FUNCTION_BLOCK DLG_CTRL (* Ablaufsteuerung eines VT-Dialogs (MessageBox) *)
  (* Standard: 61499-2; Description: Copyright (c) 2026 Meisterschulen am Ostbahnhof This program and the accompanying materials are made available under the terms of the Eclipse Public License 2.0 which is available at https://www.eclipse.org/legal/epl-2.0/ SPDX-License-Identifier: EPL-2.0 *)
  (* Version 1.0, 2026-11-17, Franz Höpfinger, Meisterschulen am Ostbahnhof, initial API and implementation and/or initial documentation *)
  PACKAGE isobus::UT::dialog;
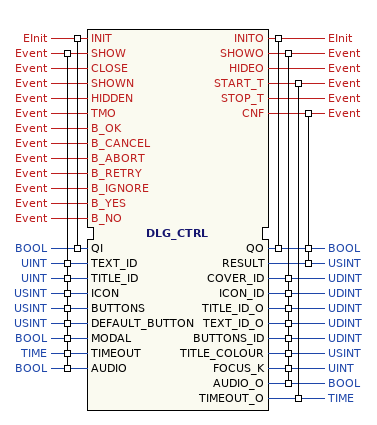
  EVENT_INPUT
    INIT : EInit WITH QI; (* Initialisierung *)
    SHOW WITH TEXT_ID, TITLE_ID, ICON, BUTTONS, DEFAULT_BUTTON, MODAL, TIMEOUT, AUDIO; (* Dialog zeigen *)
    CLOSE; (* Dialog vom Programm schliessen *)
    SHOWN; (* Anzeige-Kette fertig *)
    HIDDEN; (* Ausblenden fertig *)
    TMO; (* Zeit abgelaufen *)
    B_OK; (* Button OK losgelassen *)
    B_CANCEL; (* Button Cancel losgelassen *)
    B_ABORT; (* Button Abort losgelassen *)
    B_RETRY; (* Button Retry losgelassen *)
    B_IGNORE; (* Button Ignore losgelassen *)
    B_YES; (* Button Yes losgelassen *)
    B_NO; (* Button No losgelassen *)
  END_EVENT
  EVENT_OUTPUT
    INITO : EInit WITH QO; (* Initialisierung fertig *)
    SHOWO WITH COVER_ID, ICON_ID, TITLE_ID_O, TEXT_ID_O, BUTTONS_ID, TITLE_COLOUR, FOCUS_K, AUDIO_O; (* Anzeige-Kette starten *)
    HIDEO; (* Dialog ausblenden *)
    START_T WITH TIMEOUT_O; (* Timeout starten *)
    STOP_T; (* Timeout stoppen *)
    CNF WITH QO, RESULT; (* Dialog beendet *)
  END_EVENT
  VAR_INPUT
    QI : BOOL := TRUE; (* Freigabe *)
    TEXT_ID : UINT := UINT#65535; (* OutputString Meldungstext *)
    TITLE_ID : UINT := UINT#65535; (* OutputString Titel, NULL = Standard je Icon *)
    ICON : USINT := USINT#1; (* DLG_ICON_* *)
    BUTTONS : USINT := USINT#1; (* DLG_BTN_* *)
    DEFAULT_BUTTON : USINT := USINT#1; (* Fokus auf Taste 1..3 *)
    MODAL : BOOL := FALSE; (* Maske abdecken *)
    TIMEOUT : TIME := T#0s; (* T#0s = kein Timeout *)
    AUDIO : BOOL := FALSE; (* Ton beim Oeffnen *)
  END_VAR
  VAR_OUTPUT
    QO : BOOL; (* Qualitaet *)
    RESULT : USINT; (* DLG_RES_* *)
    COVER_ID : UDINT; (* Ziel ObjectPointer_Dlg_Cover *)
    ICON_ID : UDINT; (* Ziel ObjectPointer_Dlg_Icon *)
    TITLE_ID_O : UDINT; (* Ziel ObjectPointer_Dlg_Title *)
    TEXT_ID_O : UDINT; (* Ziel ObjectPointer_Dlg_Text *)
    BUTTONS_ID : UDINT; (* Ziel ObjectPointer_Dlg_Buttons *)
    TITLE_COLOUR : USINT; (* VT-Farbindex Titelzeile *)
    FOCUS_K : UINT; (* Fokus-Button 0..6, 7 = keiner *)
    AUDIO_O : BOOL; (* Ton ja/nein *)
    TIMEOUT_O : TIME; (* Timeout *)
  END_VAR
  VAR
    xPendingShow : BOOL; (* neues SHOW wartet *)
    xPendingClose : BOOL; (* Schliessen wartet *)
  END_VAR
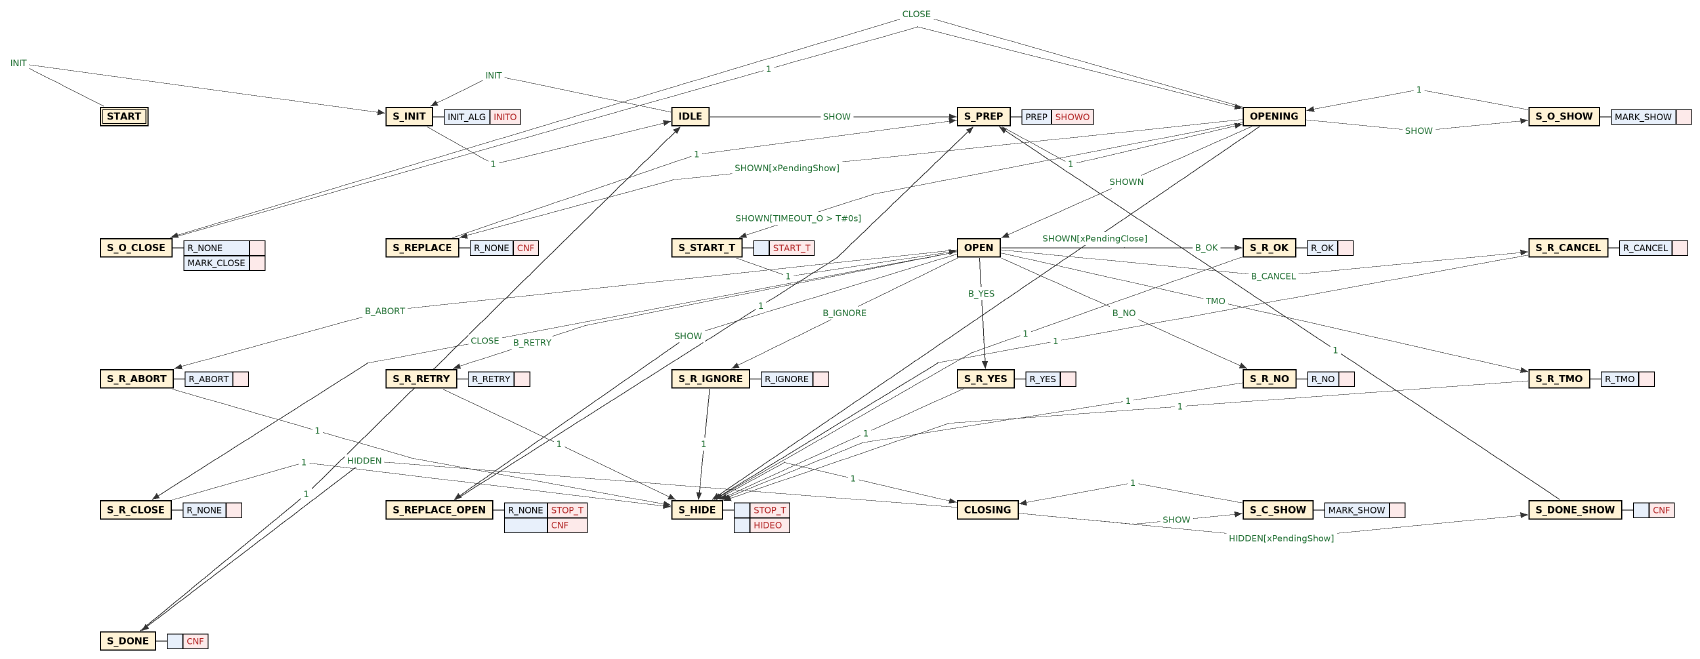
  EC_STATES
    START; (* Initial State *)
    S_INIT : INIT_ALG -> INITO;
    IDLE; (* kein Dialog offen *)
    S_PREP : PREP -> SHOWO; (* Anzeige-Kette starten *)
    OPENING; (* Anzeige-Kette laeuft *)
    S_O_SHOW : MARK_SHOW;
    S_O_CLOSE : R_NONE, MARK_CLOSE;
    S_REPLACE : R_NONE -> CNF; (* alter Dialog ersetzt *)
    S_START_T : -> START_T;
    OPEN; (* Dialog sichtbar *)
    S_R_OK : R_OK;
    S_R_CANCEL : R_CANCEL;
    S_R_ABORT : R_ABORT;
    S_R_RETRY : R_RETRY;
    S_R_IGNORE : R_IGNORE;
    S_R_YES : R_YES;
    S_R_NO : R_NO;
    S_R_TMO : R_TMO;
    S_R_CLOSE : R_NONE;
    S_REPLACE_OPEN : R_NONE -> STOP_T, -> CNF; (* neues SHOW waehrend offen *)
    S_HIDE : -> STOP_T, -> HIDEO;
    CLOSING; (* Ausblenden laeuft *)
    S_C_SHOW : MARK_SHOW;
    S_DONE_SHOW : -> CNF;
    S_DONE : -> CNF;
  END_STATES
  EC_TRANSITIONS
    START TO S_INIT := INIT;
    S_INIT TO IDLE := 1;
    IDLE TO S_INIT := INIT;
    IDLE TO S_PREP := SHOW;
    S_PREP TO OPENING := 1;
    OPENING TO S_HIDE := SHOWN[xPendingClose];
    OPENING TO S_REPLACE := SHOWN[xPendingShow];
    OPENING TO S_START_T := SHOWN[TIMEOUT_O > T#0s];
    OPENING TO OPEN := SHOWN;
    OPENING TO S_O_SHOW := SHOW;
    OPENING TO S_O_CLOSE := CLOSE;
    S_O_SHOW TO OPENING := 1;
    S_O_CLOSE TO OPENING := 1;
    S_REPLACE TO S_PREP := 1;
    S_START_T TO OPEN := 1;
    OPEN TO S_R_OK := B_OK;
    S_R_OK TO S_HIDE := 1;
    OPEN TO S_R_CANCEL := B_CANCEL;
    S_R_CANCEL TO S_HIDE := 1;
    OPEN TO S_R_ABORT := B_ABORT;
    S_R_ABORT TO S_HIDE := 1;
    OPEN TO S_R_RETRY := B_RETRY;
    S_R_RETRY TO S_HIDE := 1;
    OPEN TO S_R_IGNORE := B_IGNORE;
    S_R_IGNORE TO S_HIDE := 1;
    OPEN TO S_R_YES := B_YES;
    S_R_YES TO S_HIDE := 1;
    OPEN TO S_R_NO := B_NO;
    S_R_NO TO S_HIDE := 1;
    OPEN TO S_R_TMO := TMO;
    S_R_TMO TO S_HIDE := 1;
    OPEN TO S_R_CLOSE := CLOSE;
    S_R_CLOSE TO S_HIDE := 1;
    OPEN TO S_REPLACE_OPEN := SHOW;
    S_REPLACE_OPEN TO S_PREP := 1;
    S_HIDE TO CLOSING := 1;
    CLOSING TO S_DONE_SHOW := HIDDEN[xPendingShow];
    CLOSING TO S_DONE := HIDDEN;
    CLOSING TO S_C_SHOW := SHOW;
    S_C_SHOW TO CLOSING := 1;
    S_DONE_SHOW TO S_PREP := 1;
    S_DONE TO IDLE := 1;
  END_TRANSITIONS
  ALGORITHM INIT_ALG IN ST:
QO := QI;
RESULT := 0;
xPendingShow := FALSE;
xPendingClose := FALSE;
  END_ALGORITHM
  ALGORITHM PREP IN ST:
(* Pointer-Ziele aus der Vorlage Workspace_Dialog, IDs siehe DialogIDs.gcf *)
IF MODAL THEN COVER_ID := 14400; ELSE COVER_ID := 65535; END_IF;
CASE ICON OF
  1: ICON_ID := 3402; TITLE_COLOUR := 2;      (* gruen *)
  2: ICON_ID := 3403; TITLE_COLOUR := 15; (* navy *)
  3: ICON_ID := 3404; TITLE_COLOUR := 6;   (* oliv *)
  4: ICON_ID := 3405; TITLE_COLOUR := 12;    (* rot *)
ELSE
  ICON_ID := 65535; TITLE_COLOUR := 2;
END_CASE;
IF TITLE_ID <> 65535 THEN
  TITLE_ID_O := TITLE_ID;
ELSIF ICON >= 1 AND ICON <= 4 THEN
  TITLE_ID_O := UDINT#11409 + ICON;
ELSE
  TITLE_ID_O := 11410;
END_IF;
TEXT_ID_O := TEXT_ID;
(* FOCUS_K: 0 OK, 1 Cancel, 2 Abort, 3 Retry, 4 Ignore, 5 Yes, 6 No, 7 kein Fokus *)
FOCUS_K := 7;
CASE BUTTONS OF
  1: BUTTONS_ID := 3410; FOCUS_K := 0;
  2: BUTTONS_ID := 3411;
     IF DEFAULT_BUTTON = 2 THEN FOCUS_K := 1; ELSE FOCUS_K := 0; END_IF;
  3: BUTTONS_ID := 3412;
     IF DEFAULT_BUTTON = 2 THEN FOCUS_K := 3; ELSIF DEFAULT_BUTTON = 3 THEN FOCUS_K := 4; ELSE FOCUS_K := 2; END_IF;
  4: BUTTONS_ID := 3413;
     IF DEFAULT_BUTTON = 2 THEN FOCUS_K := 6; ELSIF DEFAULT_BUTTON = 3 THEN FOCUS_K := 1; ELSE FOCUS_K := 5; END_IF;
  5: BUTTONS_ID := 3414;
     IF DEFAULT_BUTTON = 2 THEN FOCUS_K := 6; ELSE FOCUS_K := 5; END_IF;
  6: BUTTONS_ID := 3415;
     IF DEFAULT_BUTTON = 2 THEN FOCUS_K := 1; ELSE FOCUS_K := 3; END_IF;
ELSE
  BUTTONS_ID := 65535;
END_CASE;
TIMEOUT_O := TIMEOUT;
AUDIO_O := AUDIO;
xPendingShow := FALSE;
xPendingClose := FALSE;
  END_ALGORITHM
  ALGORITHM R_NONE IN ST:
RESULT := 0;
  END_ALGORITHM
  ALGORITHM R_TMO IN ST:
RESULT := 8;
  END_ALGORITHM
  ALGORITHM MARK_SHOW IN ST:
xPendingShow := TRUE;
  END_ALGORITHM
  ALGORITHM MARK_CLOSE IN ST:
xPendingClose := TRUE;
  END_ALGORITHM
  ALGORITHM R_OK IN ST:
RESULT := 1;
  END_ALGORITHM
  ALGORITHM R_CANCEL IN ST:
RESULT := 2;
  END_ALGORITHM
  ALGORITHM R_ABORT IN ST:
RESULT := 3;
  END_ALGORITHM
  ALGORITHM R_RETRY IN ST:
RESULT := 4;
  END_ALGORITHM
  ALGORITHM R_IGNORE IN ST:
RESULT := 5;
  END_ALGORITHM
  ALGORITHM R_YES IN ST:
RESULT := 6;
  END_ALGORITHM
  ALGORITHM R_NO IN ST:
RESULT := 7;
  END_ALGORITHM
END_FUNCTION_BLOCK
